(*
SPDX-FileCopyrightText: © 2026 Oleksandr Tiutyk <trofimich@gmail.com>
SPDX-License-Identifier: MIT
License: https://opensource.org/license/mit
*)

(*!
<summary>Provides shared fixtures with early initialization for automation runner tests.</summary>
<description>
Initialized in early slot 40500 so empty sentinel arrays are available during POU variable construction.
</description>
*)

{attribute 'qualified_only'}
{attribute 'global_init_slot' := '40500'}
VAR_GLOBAL CONSTANT
	EmptyComponents : ARRAY [0..-1] OF TOF_Automation.IAutomationComponent := [];
END_VAR

(* stored: Version 1.1.0.1
   GVL AutomationRunnerTestGlobals: Id {f39300e8-8b13-4b27-bd30-9babfb0f2410} *)
